// TIA Portal project "projet_prod_offgrid" (V18)

(* hardware
DEVICE "S7-1200 station_1"  S7-1200 Station
   slot 0: "Rack_0"  S7-1200 Rack  Rack  V1.0
   slot 1: "PLC_1"  CPU 1211C DC/DC/DC  6ES7 211-1AE40-0XB0  V4.5
*)

// ===== PLC "PLC_1"  CPU 1211C DC/DC/DC =====

VAR_GLOBAL   // PLC tag table "Default tag table"
   "TEST" AT %M0.0 : Bool;
   "OKTEST" AT %Q0.1 : Bool;
   "retval www" AT %MW8 : Int;
END_VAR

TYPE "UDT_Elec_3"
   STRUCT
      U_V : Real;   // [V]
      I_A : Real;   // [A]
      P_W : Real;   // [W]
   END_STRUCT;
END_TYPE

TYPE "UDT_Battery"
   STRUCT
      SOC_Pct : Real;   // [%]
      U_V : Real;   // [V]
      P_W : Real;   // [A]
      I_A : Real;   // [W]
   END_STRUCT;
END_TYPE

TYPE "UDT_Settings"
   STRUCT
      Min_SOC_Pct : Real;
      Critical_SOC_Pct : Real;
      Gen_Enabled : Bool;
      Grid_Enabled : Bool;
      Gen_Start_Delay_s : Int;
      Parameter_Apply_Req : Bool;
      Parameter_Apply_Ack : Bool;
      Parameter_Apply_Code : Int;
      Parameter_Apply_Counter : DInt;
   END_STRUCT;
END_TYPE

TYPE "UDT_Status"
   STRUCT
      Inv_L1_1_State : Int;
      Inv_L1_1_FaultCode : Int;
      Inv_L1_2_State : Int;
      Inv_L1_2_FaultCode : Int;
      Inv_L2_1_State : Int;
      Inv_L2_1_FaultCode : Int;
      Inv_L2_2_State : Int;
      Inv_L2_2_FaultCode : Int;
      Inv_L3_1_State : Int;
      Inv_L3_1_FaultCode : Int;
      Inv_L3_2_State : Int;
      Inv_L3_2_FaultCode : Int;
      Gen_Running : Bool;
      Grid_Available : Bool;
   END_STRUCT;
END_TYPE

TYPE "UDT_AlarmSlot"
   STRUCT
      Active : Bool;
      Severity : Int;
      Source : String;
      Message : String;
      FaultCode : Int;
      Ts : DTL;
      AckReq : Bool;
      Acked : Bool;
      "Counter" : Int;
   END_STRUCT;
END_TYPE

DATA_BLOCK "DB_SCADA"   // DB1
{ S7_Optimized_Access := 'TRUE' }
VERSION : 0.1
   VAR
      Grid_L1 : "UDT_Elec_3";
      Grid_L2 : "UDT_Elec_3";
      Grid_L3 : "UDT_Elec_3";
      Grid_Freq_Hz : Real;
      PV : "UDT_Elec_3";
      Gen : "UDT_Elec_3";
      Gen_Freq_Hz : Real;
      LoadCritical_L1 : "UDT_Elec_3";
      LoadCritical_L2 : "UDT_Elec_3";
      LoadCritical_L3 : "UDT_Elec_3";
      LoadCritical_Freq_Hz : Real;
      LoadNormal : "UDT_Elec_3";
      LoadNormal_Freq_Hz : Real;
      Battery : "UDT_Battery";
      Settings : "UDT_Settings";
      Status : "UDT_Status";
      Alarms : Array[0..20] of "UDT_AlarmSlot";
      Alarms_Count : USInt := 20;
      Alarms_ActiveCount : Int;
      Alarms_CritActive : Bool;
   END_VAR
BEGIN
END_DATA_BLOCK

DATA_BLOCK "FB_Simulation_DB"   // DB2
{ S7_Optimized_Access := 'TRUE' }
VERSION : 0.1
// stored: InstanceOfName FB_Simulation
"FB_Simulation"
BEGIN
END_DATA_BLOCK

DATA_BLOCK "FB_AlarmsManager_DB"   // DB3
{ S7_Optimized_Access := 'TRUE' }
VERSION : 0.1
// stored: InstanceOfName FB_AlarmsManager
"FB_AlarmsManager"
BEGIN
END_DATA_BLOCK

DATA_BLOCK "FB_AlarmsGenerator_DB"   // DB4
{ S7_Optimized_Access := 'TRUE' }
VERSION : 0.1
// stored: InstanceOfName FB_AlarmsGenerator
"FB_AlarmsGenerator"
BEGIN
END_DATA_BLOCK

DATA_BLOCK "Parameter_Req_DB_1"   // DB5
{ S7_Optimized_Access := 'TRUE' }
VERSION : 0.1
// stored: InstanceOfName Parameter_Req
"Parameter_Req"
BEGIN
END_DATA_BLOCK

FUNCTION_BLOCK "FB_Simulation"   // FB1, SCL
{ S7_Optimized_Access := 'TRUE' }
VERSION : 0.1
   VAR
      Init_Done : Bool;
      U_Nominal : Real;
      I_Max : Real;
      dI : Real;
      dSOC : Real;
      Charge : Bool;
   END_VAR
BEGIN

   #Init_Done := FALSE;
   #U_Nominal:= 230.0;
   #I_Max:= 100.0;
   #dI := 0.5;
   #dSOC := 0.02;
   #Charge:= TRUE;

   // ================================
   // INITIALISATION (UNE SEULE FOIS)
   // ================================

   IF NOT #Init_Done THEN
       "DB_SCADA".Battery.U_V := 230.0;
       "DB_SCADA".Battery.I_A := 0.0;
       "DB_SCADA".Battery.SOC_Pct := 50.0;
       "DB_SCADA".Battery.P_W := 0.0;

       "DB_SCADA".LoadNormal.U_V := 230.0;
       "DB_SCADA".LoadNormal.I_A := 10.0;
       "DB_SCADA".LoadNormal.P_W := 2300.0;

       "DB_SCADA".LoadCritical_L1.U_V := 230.0;
       "DB_SCADA".LoadCritical_L1.I_A := 5.0;
       "DB_SCADA".LoadCritical_L1.P_W := 1150.0;

       "DB_SCADA".PV.U_V := 230.0;
       "DB_SCADA".PV.I_A := 20.0;
       "DB_SCADA".PV.P_W := 4600.0;

       "DB_SCADA".Grid_L1.U_V := 230.0;
       "DB_SCADA".Grid_L1.I_A := 0.0;
       "DB_SCADA".Grid_L1.P_W := 0.0;

       "DB_SCADA".Gen.U_V := 230.0;
       "DB_SCADA".Gen.I_A := 0.0;
       "DB_SCADA".Gen.P_W := 0.0;

       #Init_Done := TRUE;
   END_IF;


   // ================================
   // SIMULATION BATTERIE
   // ================================

   IF #Charge THEN
       "DB_SCADA".Battery.I_A := "DB_SCADA".Battery.I_A + #dI;
       "DB_SCADA".Battery.SOC_Pct := "DB_SCADA".Battery.SOC_Pct + #dSOC;
   ELSE
       "DB_SCADA".Battery.I_A := "DB_SCADA".Battery.I_A - #dI;
       "DB_SCADA".Battery.SOC_Pct := "DB_SCADA".Battery.SOC_Pct - #dSOC;
   END_IF;

   IF "DB_SCADA".Battery.SOC_Pct >= 95.0 THEN
       #Charge := FALSE;
   END_IF;

   IF "DB_SCADA".Battery.SOC_Pct <= 20.0 THEN
       #Charge := TRUE;
   END_IF;

   "DB_SCADA".Battery.P_W :=
   "DB_SCADA".Battery.U_V * "DB_SCADA".Battery.I_A;
END_FUNCTION_BLOCK

FUNCTION_BLOCK "Parameter_Req"   // FB2, SCL
{ S7_Optimized_Access := 'TRUE' }
VERSION : 0.1
   VAR
      LastCounter : DInt;
      ReqPrev : Bool;
   END_VAR
BEGIN
   #LastCounter:= -1;


   // --- READ HANDSHAKE VARS ---
   IF "DB_SCADA".Settings.Parameter_Apply_Req THEN

       // Si tu utilises le counter, on traite seulement un nouveau counter
       IF "DB_SCADA".Settings.Parameter_Apply_Counter <> #LastCounter THEN
           #LastCounter := "DB_SCADA".Settings.Parameter_Apply_Counter;

           // Par défaut OK
           "DB_SCADA".Settings.Parameter_Apply_Code := 0;

           // --- VALIDATION / CLAMP ---
           IF "DB_SCADA".Settings.Min_SOC_Pct < 0.0 THEN
               "DB_SCADA".Settings.Min_SOC_Pct := 0.0;
               "DB_SCADA".Settings.Parameter_Apply_Code := 1;
           ELSIF "DB_SCADA".Settings.Min_SOC_Pct > 100.0 THEN
               "DB_SCADA".Settings.Min_SOC_Pct := 100.0;
               "DB_SCADA".Settings.Parameter_Apply_Code := 1;
           END_IF;

           IF "DB_SCADA".Settings.Critical_SOC_Pct < 0.0 THEN
               "DB_SCADA".Settings.Critical_SOC_Pct := 0.0;
               "DB_SCADA".Settings.Parameter_Apply_Code := 1;
           ELSIF "DB_SCADA".Settings.Critical_SOC_Pct > 100.0 THEN
               "DB_SCADA".Settings.Critical_SOC_Pct := 100.0;
               "DB_SCADA".Settings.Parameter_Apply_Code := 1;
           END_IF;

           IF "DB_SCADA".Settings.Gen_Start_Delay_s < 0 THEN
               "DB_SCADA".Settings.Gen_Start_Delay_s := 0;
               "DB_SCADA".Settings.Parameter_Apply_Code := 1;
           ELSIF "DB_SCADA".Settings.Gen_Start_Delay_s > 3600 THEN
               "DB_SCADA".Settings.Gen_Start_Delay_s := 3600;
               "DB_SCADA".Settings.Parameter_Apply_Code := 1;
           END_IF;

           // --- ACK PULSE ---
           "DB_SCADA".Settings.Parameter_Apply_Ack := TRUE;

       END_IF;

   ELSE
       // Quand Req retombe, on coupe l'ACK (impulsion)
       "DB_SCADA".Settings.Parameter_Apply_Ack := FALSE;
   END_IF;
END_FUNCTION_BLOCK

FUNCTION_BLOCK "FB_AlarmsManager"   // FB3, SCL
{ S7_Optimized_Access := 'TRUE' }
VERSION : 0.1
   VAR_IN_OUT
      Alarms : Array[0..20] of "UDT_AlarmSlot";
      Alarms_ActiveCount : Int;
      Alarms_CritActive : Bool;
   END_VAR
   VAR_TEMP
      i : Int;
   END_VAR
BEGIN

   // =======================
   // 1) ACK handling
   // =======================
   FOR #i := 1 TO 20 DO
       // SCADA pulse -> Acked
       IF #Alarms[#i].AckReq THEN
           #Alarms[#i].Acked := TRUE;
           #Alarms[#i].AckReq := FALSE; // consommer le pulse (TRÈS IMPORTANT)
       END_IF;
   END_FOR;


   // =======================
   // 2) Clear policy (normal industriel)
   // =======================
   // Règle demandée : l’alarme "disparaît" quand défaut disparu ET ack.
   // -> Donc quand Active=FALSE et Acked=TRUE, on peut vider champs.
   // (Optionnel : si tu veux garder l’historique, commente cette section.)
   FOR #i := 1 TO 20 DO
       IF (NOT #Alarms[#i].Active) AND (#Alarms[#i].Acked) THEN
           // on "libère" le slot (il n’apparaîtra plus côté SCADA)
           #Alarms[#i].Severity := 0;
           #Alarms[#i].Source := '';
           #Alarms[#i].Message := '';
           #Alarms[#i].FaultCode := 0;
           // on garde Counter/Ts (ou tu peux aussi les reset si tu veux)
           // Alarms[i].Counter := 0;
           // Alarms[i].Ts := DTL#1970-01-01-00:00:00.000;
           #Alarms[#i].Acked := FALSE; // slot prêt pour prochaine alarme
       END_IF;
   END_FOR;


   // =======================
   // 3) Global counters
   // =======================
   #Alarms_ActiveCount := 0;
   #Alarms_CritActive := FALSE;

   FOR #i := 1 TO 20 DO
       IF #Alarms[#i].Active THEN
           #Alarms_ActiveCount := #Alarms_ActiveCount + 1;

           // Crit = 2 (aligné avec DB/API)
           IF #Alarms[#i].Severity = 2 THEN
               #Alarms_CritActive := TRUE;
           END_IF;
       END_IF;
   END_FOR;
END_FUNCTION_BLOCK

FUNCTION_BLOCK "FB_AlarmsGenerator"   // FB4, SCL
{ S7_Optimized_Access := 'TRUE' }
VERSION : 0.1
   VAR
      nowDTL : DTL;
      prevActive : Array[0..20] of Bool;
      "return" : Int;
   END_VAR
BEGIN

   // Helper local : déclenchement standard
   // convention : Inv_State = 3 => fault
   // severity : 0 info, 1 warn, 2 crit
   // ==============================

   // ------------------------------
   // SLOT 4 : Inverter L2-2 (ton exemple)
   // ------------------------------
   "DB_SCADA".Alarms[4].Active := ("DB_SCADA".Status.Inv_L2_2_State = 3);

   IF "DB_SCADA".Alarms[4].Active THEN
       // FRONT MONTANT => nouvelle occurrence
       IF NOT #prevActive[4] THEN
           "DB_SCADA".Alarms[4].Counter := "DB_SCADA".Alarms[4].Counter + 1;
           "DB_SCADA".Alarms[4].Acked := FALSE;
           "DB_SCADA".Alarms[4].Ts := #nowDTL;
       END_IF;

       "DB_SCADA".Alarms[4].Severity := 2; // CRIT (aligné API/DB)
       "DB_SCADA".Alarms[4].Source := 'Inv L2-2';
       "DB_SCADA".Alarms[4].Message := 'Fault detected';
       "DB_SCADA".Alarms[4].FaultCode := "DB_SCADA".Status.Inv_L2_2_FaultCode;
   END_IF;

   #prevActive[4] := "DB_SCADA".Alarms[4].Active;


   // ------------------------------
   // SLOT 1 : Inv L1-1
   // ------------------------------
   "DB_SCADA".Alarms[1].Active := ("DB_SCADA".Status.Inv_L1_1_State = 3);

   IF "DB_SCADA".Alarms[1].Active THEN
       IF NOT #prevActive[1] THEN
           "DB_SCADA".Alarms[1].Counter := "DB_SCADA".Alarms[1].Counter + 1;
           "DB_SCADA".Alarms[1].Acked := FALSE;
           "DB_SCADA".Alarms[1].Ts := #nowDTL;
       END_IF;

       "DB_SCADA".Alarms[1].Severity := 2;
       "DB_SCADA".Alarms[1].Source := 'Inv L1-1';
       "DB_SCADA".Alarms[1].Message := 'Fault detected';
       "DB_SCADA".Alarms[1].FaultCode := "DB_SCADA".Status.Inv_L1_1_FaultCode;
   END_IF;

   #prevActive[1] := "DB_SCADA".Alarms[1].Active;


   // ------------------------------
   // SLOT 2 : Inv L1-2
   // ------------------------------
   "DB_SCADA".Alarms[2].Active := ("DB_SCADA".Status.Inv_L1_2_State = 3);

   IF "DB_SCADA".Alarms[2].Active THEN
       IF NOT #prevActive[2] THEN
           "DB_SCADA".Alarms[2].Counter := "DB_SCADA".Alarms[2].Counter + 1;
           "DB_SCADA".Alarms[2].Acked := FALSE;
           "DB_SCADA".Alarms[2].Ts := #nowDTL;
       END_IF;

       "DB_SCADA".Alarms[2].Severity := 2;
       "DB_SCADA".Alarms[2].Source := 'Inv L1-2';
       "DB_SCADA".Alarms[2].Message := 'Fault detected';
       "DB_SCADA". Alarms[2].FaultCode := "DB_SCADA".Status.Inv_L1_2_FaultCode;
   END_IF;

   #prevActive[2] := "DB_SCADA".Alarms[2].Active;


   // ------------------------------
   // SLOT 3 : Inv L2-1
   // ------------------------------
   "DB_SCADA".Alarms[3].Active := ("DB_SCADA".Status.Inv_L2_1_State = 3);

   IF "DB_SCADA".Alarms[3].Active THEN
       IF NOT #prevActive[3] THEN
           "DB_SCADA".Alarms[3].Counter := "DB_SCADA".Alarms[3].Counter + 1;
           "DB_SCADA".Alarms[3].Acked := FALSE;
           "DB_SCADA".Alarms[3].Ts := #nowDTL;
       END_IF;

       "DB_SCADA".Alarms[3].Severity := 2;
       "DB_SCADA".Alarms[3].Source := 'Inv L2-1';
       "DB_SCADA".Alarms[3].Message := 'Fault detected';
       "DB_SCADA".Alarms[3].FaultCode := "DB_SCADA".Status.Inv_L2_1_FaultCode;
   END_IF;

   #prevActive[3] := "DB_SCADA".Alarms[3].Active;


   // ------------------------------
   // SLOT 5 : Inv L3-1
   // ------------------------------
   "DB_SCADA".Alarms[5].Active := ("DB_SCADA".Status.Inv_L3_1_State = 3);

   IF "DB_SCADA".Alarms[5].Active THEN
       IF NOT #prevActive[5] THEN
           "DB_SCADA".Alarms[5].Counter := "DB_SCADA".Alarms[5].Counter + 1;
           "DB_SCADA".Alarms[5].Acked := FALSE;
           "DB_SCADA".Alarms[5].Ts := #nowDTL;
       END_IF;

       "DB_SCADA".Alarms[5].Severity := 2;
       "DB_SCADA".Alarms[5].Source := 'Inv L3-1';
       "DB_SCADA".Alarms[5].Message := 'Fault detected';
       "DB_SCADA".Alarms[5].FaultCode := "DB_SCADA".Status.Inv_L3_1_FaultCode;
   END_IF;

   #prevActive[5] := "DB_SCADA".Alarms[5].Active;


   // ------------------------------
   // SLOT 6 : Inv L3-2
   // ------------------------------
   "DB_SCADA".Alarms[6].Active := ("DB_SCADA".Status.Inv_L3_2_State = 3);

   IF "DB_SCADA".Alarms[6].Active THEN
       IF NOT #prevActive[6] THEN
           "DB_SCADA".Alarms[6].Counter := "DB_SCADA".Alarms[6].Counter + 1;
           "DB_SCADA".Alarms[6].Acked := FALSE;
           "DB_SCADA".Alarms[6].Ts := #nowDTL;
       END_IF;

       "DB_SCADA".Alarms[6].Severity := 2;
       "DB_SCADA".Alarms[6].Source := 'Inv L3-2';
       "DB_SCADA".Alarms[6].Message := 'Fault detected';
       "DB_SCADA".Alarms[6].FaultCode := "DB_SCADA".Status.Inv_L3_2_FaultCode;
   END_IF;

   #prevActive[6] := "DB_SCADA".Alarms[6].Active;


   // ------------------------------
   // Exemple warning : Grid absent (slot 10)
   // ------------------------------
   "DB_SCADA".Alarms[10].Active := (NOT "DB_SCADA".Status.Grid_Available);

   IF "DB_SCADA".Alarms[10].Active THEN
       IF NOT #prevActive[10] THEN
           "DB_SCADA".Alarms[10].Counter := "DB_SCADA".Alarms[10].Counter + 1;
           "DB_SCADA".Alarms[10].Acked := FALSE;
           "DB_SCADA".Alarms[10].Ts := #nowDTL;
       END_IF;

       "DB_SCADA".Alarms[10].Severity := 1; // WARN
       "DB_SCADA".Alarms[10].Source := 'Grid';
       "DB_SCADA".Alarms[10].Message := 'Grid not available';
       "DB_SCADA".Alarms[10].FaultCode := 0;
   END_IF;

   #prevActive[10] := "DB_SCADA".Alarms[10].Active;
END_FUNCTION_BLOCK

ORGANIZATION_BLOCK "Main"   // OB1, LAD, ProgramCycle
TITLE = "Main Program Sweep (Cycle)"
{ S7_Optimized_Access := 'TRUE' }
VERSION : 0.1
   VAR_INPUT
      Initial_Call : Bool;   // Initial call of this OB
      Remanence : Bool;   // =True, if remanent data are available
   END_VAR
BEGIN

REGION Network 1
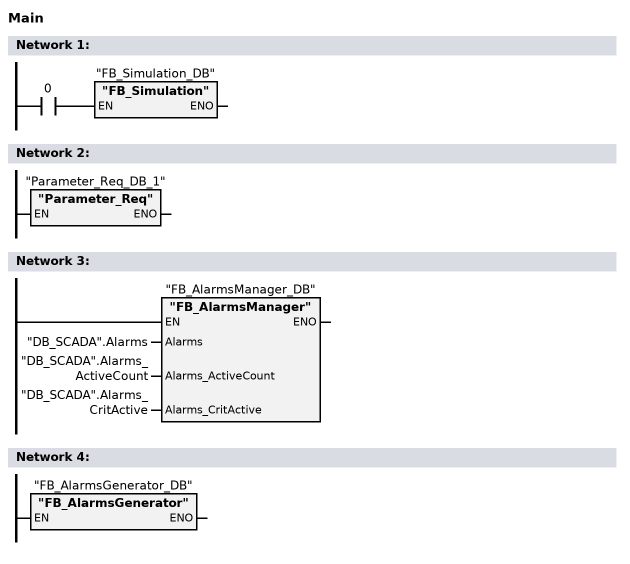
   RUNG wire#powerrail
      Contact( 0 )
      "FB_Simulation_DB"()
   END_RUNG
   // the same network as SCL:
   IF 0 THEN
       "FB_Simulation_DB"();   // "FB_Simulation"
   END_IF;
END_REGION

REGION Network 2
   RUNG wire#powerrail
      "Parameter_Req_DB_1"()
   END_RUNG
   // the same network as SCL:
   "Parameter_Req_DB_1"();   // "Parameter_Req"
END_REGION

REGION Network 3
   RUNG wire#powerrail
      "FB_AlarmsManager_DB"(Alarms := "DB_SCADA".Alarms, Alarms_ActiveCount := "DB_SCADA".Alarms_ActiveCount, Alarms_CritActive := "DB_SCADA".Alarms_CritActive)
   END_RUNG
   // the same network as SCL:
   "FB_AlarmsManager_DB"(Alarms := "DB_SCADA".Alarms,   // "FB_AlarmsManager"
                         Alarms_ActiveCount := "DB_SCADA".Alarms_ActiveCount,
                         Alarms_CritActive := "DB_SCADA".Alarms_CritActive);
END_REGION

REGION Network 4
   RUNG wire#powerrail
      "FB_AlarmsGenerator_DB"()
   END_RUNG
   // the same network as SCL:
   "FB_AlarmsGenerator_DB"();   // "FB_AlarmsGenerator"
END_REGION
END_ORGANIZATION_BLOCK